(*
SPDX-FileCopyrightText: c 2026 Oleksandr Tiutyk <trofimich@gmail.com>
SPDX-License-Identifier: MIT
License: https://opensource.org/license/mit
*)

(*!
<summary>Checks full and windowed joining and cursor reuse after insufficient capacity.</summary>
<description>
Uses one task and stays at a stable address while assertions are bound to this instance.
</description>
*)

{attribute 'no_assign'}
{attribute 'no_explicit_call' := 'do not call this function block directly'}
FUNCTION_BLOCK WideStringJoinTest EXTENDS TOF_Testing.SingleCycleTest
VAR_STAT
	{attribute 'hide'}
	_ClassName : STRING := __POUNAME();
END_VAR
VAR
	_Source : WSTRING := "123 , , 456, 789 ,0";
	_Splitter : TOF_Core.WideStringSplittingEnumerator;
END_VAR

(*!
<summary>Checks full and windowed joining and cursor reuse after insufficient capacity.</summary>
<description>
Owns a persistent cursor and its borrowed source. Reset releases the current fragment before the result is reported.
</description>
*)
METHOD PROTECTED ExecuteTest
VAR
	separator : WSTRING := ",";
	joined : WSTRING := "old target";
	shortTarget : WSTRING(2);
	accepted : BOOL;
END_VAR
_Splitter := TOF_Core.WideStrings.CreateSplitter(sourceString := _Source, separator := separator);
TOF_Core.WideStrings.Join(targetString := joined, separator := separator, sourceEnumerator := _Splitter);
Assert.ThatBool(
	actual := joined = _Source,
	message := "Unrestricted Join must reconstruct all fragments including their whitespace"
).IsTrue();

_Splitter.Reset();
_Splitter := TOF_Core.WideStrings.CreateSplitter(
	sourceString := _Source,
	separator := separator,
	maxCount := 3,
	trimEntries := TRUE,
	removeEmptyEntries := TRUE
);
TOF_Core.WideStrings.Join(
	targetString := joined,
	separator := separator,
	sourceEnumerator := _Splitter,
	startIndex := 1,
	count := 2
);
Assert.ThatBool(
	actual := joined = "456,789",
	message := "The requested window must contain fragments 1 and 2"
).IsTrue();

_Splitter.Reset();
accepted := TOF_Core.WideStrings.TryJoin(targetString := shortTarget, separator := separator, sourceEnumerator := _Splitter);
Assert.ThatBool(
	actual := accepted,
	message := "TryJoin must reject a target too small for the first fragment"
).IsFalse();

_Splitter.Reset();
accepted := TOF_Core.WideStrings.TryJoin(
	targetString := joined,
	separator := separator,
	sourceEnumerator := _Splitter,
	count := 1
);
Assert.ThatBool(
	actual := accepted AND_THEN joined = "123",
	message := "After Reset, TryJoin must restart and replace the old target text"
).IsTrue();
END_METHOD

(*!
<summary>Resets the splitter and releases any active fragment before reporting.</summary>
<description>
Safe after partial initialization and after explicit cleanup in the scenario.
</description>
*)
METHOD PROTECTED AfterTest
_Splitter.Reset();
END_METHOD

//! <summary>Borrows the concrete class name. Callers must not modify it.</summary>
{attribute 'monitoring' := 'call'}
PROPERTY ClassName : REFERENCE TO STRING
GET
ClassName REF= _ClassName;
END_GET
END_PROPERTY

//! <summary>Borrows the compiler-initialized namespace name. Callers must not modify it.</summary>
{attribute 'monitoring' := 'call'}
PROPERTY NamespaceName : REFERENCE TO STRING
GET
NamespaceName REF= CurrentNamespace.Name;
END_GET
END_PROPERTY

//! <summary>Reports the concrete instance size in bytes.</summary>
{attribute 'monitoring' := 'call'}
PROPERTY SelfSize : ULINT
GET
SelfSize := XSIZEOF(THIS^);
END_GET
END_PROPERTY

END_FUNCTION_BLOCK

(* stored: Version 1.1.0.1
   POU WideStringJoinTest: Id {e49ea7c4-ece1-43cc-aa2b-0bb7ffdd8ff9}, SpecialFunc None
   Method ExecuteTest: Id {9a6cfb95-5e59-43db-beec-1530becc1239}
   Method AfterTest: Id {238721c5-7646-4a36-bd0b-2e43a14561d5}
   Property ClassName: Id {5ff5b395-2005-4d17-931f-67bd7e973ced}
   Get Get: Id {ef8fa447-2242-4f69-8e3f-306efb0b4bd5}
   Property NamespaceName: Id {5af7da0c-100b-4595-ae5e-02b979d1593b}
   Get Get: Id {5b4e6766-7083-4441-8cde-c521326c7005}
   Property SelfSize: Id {73ebb43d-700a-4210-94d4-218e2bf86114}
   Get Get: Id {423e0c0c-3131-470c-8a61-55bb24ef7660} *)
